PROGRAM Rs232Logging
VAR


	fbPcCom		: FB_SerialCom;
	
	(* exchange buffers with background communication with the PC COM port device *)
	RxBufferPcCom	: ComBuffer;	(* Receive data buffer; used with all receive function blocks *)
	TxBufferPcCom	: ComBuffer;	(* Transmit data buffer; used with all receive function blocks *)
	
END_VAR

VAR_OUTPUT
	rWeight: REAL;
END_VAR




(* background communication with the PC COM port device *)
BackgroundPcCOM(RxBufferPcCom:=RxBufferPcCom, TxBufferPcCom:=TxBufferPcCom);


(* Send and receive commands *)
fbPcCom(TxBuffer:=TxBufferPcCom, RxBuffer:=RxBufferPcCom);
	
 rWeight:=fbPcCom.Weight;

END_PROGRAM

(* stored: Version 1.1.0.1, ProductVersion 3.1.4024.12
   POU Rs232Logging: Id {bc424776-4580-4a06-af9d-303a952ea526}, SpecialFunc None *)
